// TIA Portal V21 export
// export: Created 2026-11-10T07:02:22.6088582Z, ExportSetting WithDefaults, DisplayName Totally Integrated Automation Portal, DisplayVersion V21 Update 3, DisplayName STEP 7 Professional, DisplayVersion V21 Update 3, DisplayName STEP 7 Safety, DisplayVersion V21, DisplayName Tech WebApplication, DisplayVersion V21, DisplayName WinCC Basic/Comfort/Advanced, DisplayVersion V21 Update 3, DisplayName WinCC Unified, DisplayVersion V21 Update 3
FUNCTION_BLOCK "FB_SclCalls"   // FB3, SCL
{ S7_Optimized_Access := 'TRUE' }
VERSION : 0.1
// stored: AutoNumber true, IsIECCheckEnabled false, IsRetainMemResEnabled false, MemoryReserve 100, SetENOAutomatically false, UDAEnableTagReadback false
   VAR_INPUT
      start : Bool;
      pt : Time;
   END_VAR
   VAR_OUTPUT
      q : Bool;
      cnt : Int;
   END_VAR
   VAR
      tonInst { S7_SetPoint := 'True'} : TON_TIME;
      tofInst { S7_SetPoint := 'True'} : TOF_TIME;
      tpInst { S7_SetPoint := 'True'} : TP_TIME;
      ctuInst { S7_SetPoint := 'True'} : CTU_INT;
      trig { S7_SetPoint := 'True'} : R_TRIG;
      ftrig { S7_SetPoint := 'True'} : F_TRIG;
      "counter" : Int;
      ifc { S7_SetPoint := 'True'} : "FB_Iface";
   END_VAR
   VAR_TEMP
      r : Real;
      "b" : Bool;
      res : Int;
      tot : Int;
   END_VAR
BEGIN
   #tonInst(IN := #start, PT := #pt);
   #q := #tonInst.Q;
   #tofInst(IN := #start, PT := T#2s);
   #tpInst(IN := #start, PT := #pt, Q => #b);
   #ctuInst(CU := #start, R := FALSE, PV := 10);
   #cnt := #ctuInst.CV;
   #trig(CLK := #start);
   IF #trig.Q THEN
       #counter := 0;
   END_IF;
   #ftrig(CLK := #start);
   #b := #ftrig.Q;
   #ifc(iBool := TRUE, iInt := 2, iReal := 1.0, ioReal := #r);
   #cnt := #ifc.oInt;
   "FB_Iface_DB"(iBool := #start, iInt := #cnt, iReal := #r, ioReal := #r, oInt => #cnt);
   "FC_SclOps"();
   #res := "FC_SclCtl"(n := 5, flag := TRUE, total => #tot);
   #res := "FC_SclCtl"(n := #res, flag := #b, total => #tot);
END_FUNCTION_BLOCK
